(* IEC 61131-3 sources: StructuredFuzzer/code_analysis/src/programs/depth/depth_1, 1 file *)

(* ---- depth_1.st ---- *)
PROGRAM My_Program
  VAR
    button1 AT %IX0.0 : BOOL := FALSE;
    led AT %QX0.0 : BOOL;
  END_VAR

  IF button1 = TRUE THEN
    led := TRUE;
  ELSE
    led := FALSE;
  END_IF;
END_PROGRAM

CONFIGURATION STD_CONF

  RESOURCE STD_RESSOURCE ON PLC
    TASK TaskMain(INTERVAL := T#50ms,PRIORITY := 0);
    PROGRAM Inst0 WITH TaskMain : My_Program;
  END_RESOURCE
END_CONFIGURATION
